NAMESPACE TiaMcp_UnitA
TYPE "TiaMcpComponentState"
VERSION : 0.1
STRUCT
    Active : Bool;
END_STRUCT;
END_TYPE
END_NAMESPACE
